// TIA Portal V20 export
TYPE "T_CON_DATA"
   STRUCT
      TCON : Struct
         IN : Struct
            START : Bool;
            ID : CONN_OUC;
         END_STRUCT;
         OUT : Struct
            DONE : Bool;
            BYSY : Bool;
            ERROR : Bool;
            STATUS : Word;
         END_STRUCT;
      END_STRUCT;
   END_STRUCT;
END_TYPE
